// TIA Portal V20 export
TagTable "Plant tags"
  Motor_1_Run :   (500 ms)
  Motor_2_Run :   (1 s)
